Staubli VAL3: Force6Item.dtx

mdesc mNomSpeed
public string sArmType
public num nMaxJnt6Force[6]
